Fanuc KAREL source: KT00795.KL

PROGRAM KT00795
%NOLOCKGROUP
VAR
  S1: STRING[80]
  S2: STRING[80]
  OUT: REAL
BEGIN
  S1 = 'A'
  S2 = 'B'
  S1 = 'A'
  S2 = 'B'
  OUT = COS(S1)
END KT00795
